Staubli VAL3: start.pgx

program start()
begin
  taskCreate "appMain",20,Main()
end
